(* IEC 61131-3 sources: codesys-to-s7/tests/corpus/C2S7-ADDR-OVERLAP/neg, 1 file *)

(* ---- input.st ---- *)
VAR_GLOBAL
    wA AT %MW5 : WORD;
    iA AT %MW5 : INT;
END_VAR
